DATA_BLOCK "GDB_GRAPH_PressDemoHome"
{ S7_Optimized_Access := 'TRUE' }
VERSION : 0.1
NON_RETAIN
"FB_GRAPH_PressDemoHome"
BEGIN
END_DATA_BLOCK
